Fanuc KAREL source: ko00037.KL

-- PROVISIONAL review KL for V770-1; original PC SHA256 a50fb7aecdb75a4a7877a812d204d3d2a256b28427c3476117e1ef6a1ad8d7aa
-- Incomplete behavior may be omitted. Consult companion uncertainty JSON. Do not deploy.
PROGRAM KO00037
%NOLOCKGROUP
BEGIN
  -- UNRESOLVED_PC offsets 5-12; opcodes 9D,23
  -- UNRESOLVED_PC offsets 17-69; opcodes 27,27,49,7E,AD,27,49,7E,AD,22,31,7E,4A
  -- UNRESOLVED_PC offsets 74-78; opcodes 7F
END KO00037
